// TIA Portal V21 export
// export: Created 2026-11-08T20:57:50.8689948Z, ExportSetting WithDefaults, DisplayName Totally Integrated Automation Portal, DisplayVersion V21 Update 3, DisplayName STEP 7 Professional, DisplayVersion V21 Update 3, DisplayName STEP 7 Safety, DisplayVersion V21, DisplayName Tech WebApplication, DisplayVersion V21, DisplayName WinCC Basic/Comfort/Advanced, DisplayVersion V21 Update 3, DisplayName WinCC Unified, DisplayVersion V21 Update 3
FUNCTION "FC_Stl" : Void   // FC1, STL
TITLE = STL test FC
{ S7_Optimized_Access := 'TRUE' }
VERSION : 0.1
// stored: AutoNumber true, UDAEnableTagReadback false
   VAR_INPUT
      "a" : Bool;
      "b" : Bool;
      x : Int;
      y : Int;
   END_VAR
   VAR_OUTPUT
      q : Bool;
      sum : Int;
   END_VAR
   VAR_TEMP
      t : Int;
   END_VAR
BEGIN

NETWORK
TITLE = Bit logic
// Network comment line 1
      A     #"a";  // and a
      AN    #"b";
      =     #q;

NETWORK
TITLE = Arithmetic
      L     #x;
      L     #y;
      +I;
      T     #t;

      L     #t;
      L     0;
      >I;
      JC    M001;
      L     0;
      T     #t;
M001: L     #t;
      T     #sum;
END_FUNCTION
